Staubli VAL3: main.pgx

program main()
begin
  close(tCurrentTool)
  pPointRs.config.shoulder = lefty
  pPointRs2.config.shoulder = lefty
  mCurrentSpeed.tvel = 100.00
  mCurrentSpeed.blend = joint
  mCurrentSpeed.reach = 0.010
  mCurrentSpeed.leave = 0.010
  // Program SpeedProg start
  // Program generated by RoboDK v6.0.7 for Staubli TS20 FL 100 TC on XX/XX/XXXX 18:00:00
  // Using nominal kinematics.
  mCurrentSpeed.reach = 0.300
  mCurrentSpeed.leave = 0.300
  mCurrentSpeed.tvel = 1.000
  call MoveLine(-607.850,543.849,363.215,136.262,30.757,-130.375)
  call MoveJoint(10.00000,-20.00000,50.00000,30.00000)
  mCurrentSpeed.reach = 1.000
  mCurrentSpeed.leave = 1.000
  mCurrentSpeed.tvel = 12.300
  call MoveLine(-640.584,506.980,371.534,136.262,30.757,-130.375)
  call MoveJoint(30.00000,25.00000,80.00000,-45.00000)
  mCurrentSpeed.reach = 2.500
  mCurrentSpeed.leave = 2.500
  mCurrentSpeed.tvel = 99.900
  call MoveLine(-607.850,543.849,363.215,136.262,30.757,-130.375)
  call MoveJoint(10.00000,-20.00000,50.00000,30.00000)
  mCurrentSpeed.reach = 3.700
  mCurrentSpeed.leave = 3.700
  mCurrentSpeed.tvel = 333.333
  call MoveLine(-640.584,506.980,371.534,136.262,30.757,-130.375)
  call MoveJoint(30.00000,25.00000,80.00000,-45.00000)
  mCurrentSpeed.reach = 6.000
  mCurrentSpeed.leave = 6.000
  mCurrentSpeed.tvel = 1000.000
  call MoveLine(-607.850,543.849,363.215,136.262,30.757,-130.375)
  call MoveJoint(10.00000,-20.00000,50.00000,30.00000)
  mCurrentSpeed.reach = 9.000
  mCurrentSpeed.leave = 9.000
  mCurrentSpeed.tvel = 2500.000
  call MoveLine(-640.584,506.980,371.534,136.262,30.757,-130.375)
  call MoveJoint(30.00000,25.00000,80.00000,-45.00000)
  mCurrentSpeed.reach = 15.000
  mCurrentSpeed.leave = 15.000
  mCurrentSpeed.tvel = 5000.000
  call MoveLine(-607.850,543.849,363.215,136.262,30.757,-130.375)
  call MoveJoint(10.00000,-20.00000,50.00000,30.00000)
  mCurrentSpeed.reach = 30.000
  mCurrentSpeed.leave = 30.000
  mCurrentSpeed.tvel = 12000.000
  call MoveLine(-640.584,506.980,371.534,136.262,30.757,-130.375)
  call MoveJoint(30.00000,25.00000,80.00000,-45.00000)
  mCurrentSpeed.reach = 75.000
  mCurrentSpeed.leave = 75.000
  mCurrentSpeed.tvel = 0.500
  call MoveLine(-607.850,543.849,363.215,136.262,30.757,-130.375)
  call MoveJoint(10.00000,-20.00000,50.00000,30.00000)
  mCurrentSpeed.reach = 150.000
  mCurrentSpeed.leave = 150.000
  mCurrentSpeed.tvel = 750.000
  call MoveLine(-640.584,506.980,371.534,136.262,30.757,-130.375)
  call MoveJoint(30.00000,25.00000,80.00000,-45.00000)
  call MoveLine(-640.584,506.980,371.534,136.262,30.757,-130.375)

  waitEndMove()
  // Program SpeedProg end

end
